(* PLC project codesys-P5-langmatrix-app.project, CODESYS CODESYS V3.5 SP17 Patch 3 *)
(* stored: creationDateTime 2026-10-20T02:17:13.2234347, modificationDateTime 1601-01-01T03:00:00 *)

// lang-matrix: ST
PROGRAM PRG_LangSt
VAR
    xA : BOOL;
    xB : BOOL;
    xQ : BOOL;
    xDone : BOOL;
    iLevel : INT;
    xHigh : BOOL;
    wCode : WORD;
    sHex : STRING;
    fbTon : TON;
    fbHyst : HYSTERESIS;
END_VAR

                  // Standard: TON; Util: HYSTERESIS; блок под замену: OSU.WORD_TO_HEX_STR (OwenStringUtils)
xQ := xA AND xB;
fbTon(IN := xQ, PT := T#100MS);
xDone := fbTon.Q;
fbHyst(IN := iLevel, HIGH := 80, LOW := 20, OUT => xHigh);
sHex := OSU.WORD_TO_HEX_STR(wInput := wCode, xUpperCase := TRUE, sPrefix := '0x');

                
END_PROGRAM

// lang-matrix: FBD
PROGRAM PRG_LangFbd
VAR
    xA : BOOL;
    xB : BOOL;
    xQ : BOOL;
    xDone : BOOL;
    iLevel : INT;
    xHigh : BOOL;
    wCode : WORD;
    sHex : STRING;
    fbTon : TON;
    fbHyst : HYSTERESIS;
END_VAR

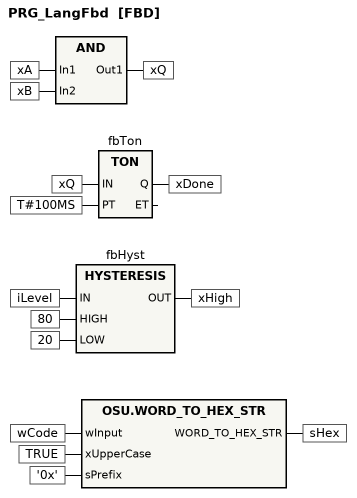
(* FBD diagram, written out as Structured Text *)
xQ := xA AND xB;
fbTon(IN := xQ, PT := T#100MS);
xDone := fbTon.Q;
fbHyst(IN := iLevel, HIGH := 80, LOW := 20);
xHigh := fbHyst.OUT;
sHex := OSU.WORD_TO_HEX_STR(wCode, TRUE, '0x');
END_PROGRAM

// lang-matrix: LD
PROGRAM PRG_LangLd
VAR
    xA : BOOL;
    xB : BOOL;
    xQ : BOOL;
END_VAR

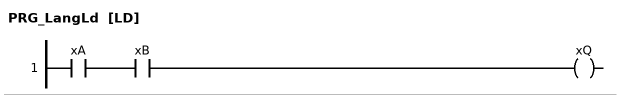
(* LD diagram, written out as Structured Text *)

xQ := xA AND xB;
END_PROGRAM

// lang-matrix: CFC
PROGRAM PRG_LangCfc
VAR
    xA : BOOL;
    xB : BOOL;
    xQ : BOOL;
    xDone : BOOL;
    iLevel : INT;
    xHigh : BOOL;
    wCode : WORD;
    sHex : STRING;
    fbTon : TON;
    fbHyst : HYSTERESIS;
END_VAR

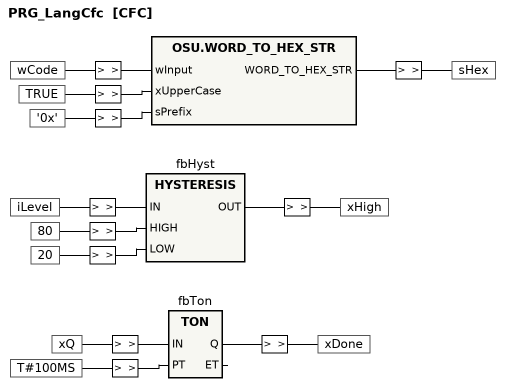
(* CFC diagram, written out as Structured Text *)
fbTon(IN := xQ, PT := T#100MS);
xDone := fbTon.Q;
fbHyst(IN := iLevel, HIGH := 80, LOW := 20);
xHigh := fbHyst.OUT;
sHex := OSU.WORD_TO_HEX_STR(wCode, TRUE, '0x');
END_PROGRAM

// lang-matrix: SFC
PROGRAM PRG_LangSfc
VAR
    xA : BOOL;
    xB : BOOL;
    xQ : BOOL;
    xDone : BOOL;
    iLevel : INT;
    xHigh : BOOL;
    wCode : WORD;
    sHex : STRING;
    fbTon : TON;
    fbHyst : HYSTERESIS;
END_VAR

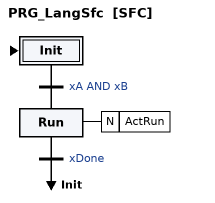
INITIAL_STEP Init:
END_STEP
TRANSITION FROM Init TO Run
  := xA AND xB;
END_TRANSITION
STEP Run:
  ActRun(N);
END_STEP
TRANSITION FROM Run TO Init
  := xDone;
END_TRANSITION

ACTION ActRun:
                      fbTon(IN := TRUE, PT := T#100MS);
xDone := fbTon.Q;
fbHyst(IN := iLevel, HIGH := 80, LOW := 20, OUT => xHigh);
sHex := OSU.WORD_TO_HEX_STR(wInput := wCode, xUpperCase := TRUE, sPrefix := '0x');

                    
END_ACTION
END_PROGRAM

// lang-matrix: вызов всех POU
PROGRAM PRG_LangMain
VAR
END_VAR

                  // Вызов POU всех языков матрицы
PRG_LangSt();
PRG_LangFbd();
PRG_LangLd();
PRG_LangCfc();
PRG_LangSfc();
PRG_LangIl();

                
END_PROGRAM
